(* IEC 61131-3 sources: canworks/test/plc_modbus, 6 files *)

(* ---- bridge_model.st ---- *)
(*
 * The bridge's control block and SDO registers for the block tests
 * (test/plc_modbus/run.sh), working on the blocks' LINK words directly
 * (library/modbus: 0-3 status, 4-6 control, 7-13 SDO request, 14-20 SDO
 * response): one call is one Modbus poll round. Mirrors ControlBlock and
 * SdoBridgeRegisters in plugin/src/bridge/bridge_blocks.cpp: a request runs
 * when its counter changes, the response echoes the counter. A read answers
 * 16#123456nn (nn the node); SILENT_NODE stays busy, ABORT_NODE aborts with
 * 16#06020000, writes without ALLOW_WRITE abort with 16#08000020;
 * RESTARTED answers as a bridge that just started with the request in place
 * (control result 6, SDO abort 16#08000021).
 * STruC++'s test runner does not copy a source block's in-out back, so a
 * test writes `link := bridge.LINK;` after each call.
 *)
FUNCTION_BLOCK BridgeModel
VAR_INPUT
  ALLOW_WRITE : BOOL := TRUE;
  SILENT_NODE : USINT := 99;
  ABORT_NODE : USINT := 98;
  REFUSE : BOOL;
  RESTARTED : BOOL;
END_VAR
VAR_OUTPUT
  LAST_CMD : WORD;
  LAST_NET : WORD;
  LAST_NODE : WORD;
  WRITTEN : UDINT;
  WRITTEN_SIZE : WORD;
  REQUESTS : INT;
  CONTROLS : INT;
END_VAR
VAR_IN_OUT
  LINK : ARRAY[0..1279] OF WORD;
END_VAR
VAR
  cmd : WORD;
  node : WORD;
END_VAR
  IF LINK[4] <> LINK[2] THEN
    LINK[2] := LINK[4];
    CONTROLS := CONTROLS + 1;
    LAST_CMD := SHR(LINK[5], 8);
    LAST_NET := LINK[5] AND 16#00FF;
    LAST_NODE := SHR(LINK[6], 8);
    IF RESTARTED THEN
      LINK[3] := 16#0600;
    ELSIF REFUSE THEN
      LINK[3] := 16#0500;
    ELSIF LAST_NET > 0 THEN
      LINK[3] := 16#0200;
    ELSE
      LINK[3] := 0;
    END_IF;
  END_IF;
  IF LINK[7] <> LINK[14] THEN
    LINK[14] := LINK[7];
    REQUESTS := REQUESTS + 1;
    cmd := SHR(LINK[8], 8);
    node := SHR(LINK[9], 8);
    LINK[16] := 0;
    LINK[17] := 0;
    LINK[18] := 0;
    LINK[19] := 0;
    IF RESTARTED THEN
      LINK[15] := 16#0300;
      LINK[16] := 16#0800;
      LINK[17] := 16#0021;
    ELSIF cmd = 2 AND NOT ALLOW_WRITE THEN
      LINK[15] := 16#0300;
      LINK[16] := 16#0800;
      LINK[17] := 16#0020;
    ELSIF node = USINT_TO_WORD(SILENT_NODE) THEN
      LINK[15] := 16#0100;
    ELSIF node = USINT_TO_WORD(ABORT_NODE) THEN
      LINK[15] := 16#0300;
      LINK[16] := 16#0602;
    ELSE
      LINK[15] := 16#0200;
      IF cmd = 1 THEN
        LINK[18] := 16#1234;
        LINK[19] := 16#5600 OR node;
      ELSE
        WRITTEN := DWORD_TO_UDINT(SHL(WORD_TO_DWORD(LINK[12]), 16) OR WORD_TO_DWORD(LINK[13]));
        WRITTEN_SIZE := SHR(LINK[11], 8);
      END_IF;
    END_IF;
  END_IF;
END_FUNCTION_BLOCK

(* ---- mailbox_model.st ---- *)
(*
 * The bridge's mailboxes for the block tests (test/plc_modbus/run.sh),
 * working on the blocks' LINK words directly (the places CW_LINK_SERVICE
 * describes): one call is one Modbus poll round of the bridge. Mirrors
 * plugin/src/bridge/mailboxes.cpp: a request runs when its counter changes
 * (an operation answers busy for one round, then done), the response echoes
 * the counter; STAGE and FETCH move data in 128-byte parts; receivers get
 * records in batches the program acknowledges; info and the cyclic table
 * are refreshed every round. Networks 0 and 1 exist. The bus is a set of
 * fixed answers:
 *   SDO node 98 aborts with 16#06020000, node 99 times out (2); 0x1008 the
 *   text "Valve block 24 V", 0x2000 600 bytes (byte i = i MOD 251), 0x2001
 *   300 bytes 'A' without a NUL, 0x6000 REAL32 1.5, 0x6001 REAL64 -2.25,
 *   0x6002 5 bytes, any other 16#12345600 + node (4 bytes);
 *   J1939 requests: PGN 65282 answers 40 bytes (i + 1), 65000 300 bytes
 *   (i MOD 256), 59999 a NACK (12, ACK_CODE 1), others 8 bytes (i);
 *   DM1/DM2 of any source but 77 (13): lamps 16#44, flash 16#04, codes
 *   16#00012304 and 16#0005A1FF, age 1500 ms;
 *   FIND_ECU knows one ECU, NAME 16#A00000000000ABCD at 16#33.
 * Messages come in with INJ_CAN, INJ_J1939, INJ_EMCY (INJ_RESTART: a new
 * CANopen session record); HOLD keeps them waiting for one batch; CLOSE_SLOT
 * closes a receiver as a stall would.
 * STruC++'s test runner does not copy a source block's in-out back, so a
 * test writes `link := bridge.LINK;` after each call.
 *)
FUNCTION_BLOCK MailboxModel
VAR_INPUT
  INJ_CAN : BOOL;
  INJ_J1939 : BOOL;
  INJ_EMCY : BOOL;
  INJ_RESTART : BOOL;
  INJ_ID : UDINT;
  INJ_EXT : BOOL;
  INJ_DLC : USINT := 8;
  INJ_LEN : UINT := 8;
  INJ_SRC : USINT;
  INJ_NODE : USINT;
  INJ_CODE : WORD;
  INJ_B0 : BYTE;
  CLOSE_SLOT : INT := -1;
  NO_J1939 : BOOL;
  HOLD : BOOL;           (* no new batch this round *)
  SKIP_MS : WORD;        (* extra milliseconds on the bridge's clock this round *)
  RX_BLOCKS : INT := 1;  (* receive_blocks: 95 record words, 215 with 2 *)
END_VAR
VAR_OUTPUT
  TX_COUNT : INT;
  TX_ID : UDINT;
  TX_DLC : WORD;
  TX_FLAGS : WORD;
  TX_B0 : BYTE;
  STAGES : INT;
  FETCHES : INT;
  REQUESTS : INT;
  W_LEN : UINT;
  W_KIND : WORD;
  W_SIZE : WORD;
  W_INDEX : WORD;
  J_PGN : UDINT;
  J_DEST : WORD;
  J_PRIO : WORD;
  J_LEN : UINT;
  J_COUNT : INT;
  DM_CLEARED : WORD;
  CYC_SETS : INT;
  CYC_STOPS : INT;
  STALLS : INT;
  OPEN_RX : INT;
END_VAR
VAR_IN_OUT
  LINK : ARRAY[0..1279] OF WORD;
END_VAR
VAR
  tick : WORD := 16#1000;
  seen : ARRAY[0..3] OF WORD;
  busy : ARRAY[0..3] OF INT;      (* rounds left before a running operation ends *)
  staged : ARRAY[0..7139] OF BYTE;
  staged_len : ARRAY[0..3] OF UINT;
  result : ARRAY[0..7139] OF BYTE;
  result_len : ARRAY[0..3] OF UINT;
  w_data : ARRAY[0..1784] OF BYTE;
  j_data : ARRAY[0..1784] OF BYTE;
  r : ARRAY[0..23] OF WORD;          (* results of the 4 mailboxes, 6 each *)
  st : ARRAY[0..3] OF WORD;          (* state << 8 | error *)
  rx_on : ARRAY[0..31] OF BOOL;
  rx_kind : ARRAY[0..31] OF WORD;
  rx_id : ARRAY[0..31] OF UDINT;
  rx_mask : ARRAY[0..31] OF UDINT;
  rx_flags : ARRAY[0..31] OF WORD;
  rx_gen : ARRAY[0..31] OF WORD;
  rx_drop : ARRAY[0..31] OF WORD;
  next_gen : WORD := 1;
  held : ARRAY[0..1784] OF BYTE;
  held_len : UINT;
  held_slot : INT := -1;
  (* Waiting records: receiver, kind, id/PGN/node, length, first byte, source, code, flags. *)
  q_n : INT;
  q_slot : ARRAY[0..63] OF INT;
  q_kind : ARRAY[0..63] OF WORD;
  q_id : ARRAY[0..63] OF UDINT;
  q_len : ARRAY[0..63] OF UINT;
  q_b0 : ARRAY[0..63] OF BYTE;
  q_src : ARRAY[0..63] OF WORD;
  q_code : ARRAY[0..63] OF WORD;
  q_flags : ARRAY[0..63] OF WORD;
  q_ext : ARRAY[0..63] OF BOOL;
  seq : WORD := 16#4000;
  present : DWORD;
  used : INT;
  acked : BOOL := TRUE;
  shown_rounds : INT;
  words : ARRAY[0..214] OF WORD;
  job_on : ARRAY[0..15] OF BOOL;
  job_gen : ARRAY[0..15] OF WORD;
  job_count : ARRAY[0..15] OF UDINT;
  job_keep : ARRAY[0..15] OF WORD;
  job_idle : ARRAY[0..15] OF INT;
  job_data : ARRAY[0..15] OF WORD;
  info_count : WORD;
  m : INT;
  n : INT;
  i : INT;
  k : INT;
  b : INT;
  op : WORD;
  net : WORD;
  len : UINT;
  slot : INT;
  jobs : INT;
  pending : DWORD;
  taken_long : DWORD;
  size : INT;
  room : BOOL;
  batch_tick : WORD;     (* the batch time's low word *)
  bits : DWORD;
END_VAR
  tick := tick + 10 + SKIP_MS;
  n := WORD_TO_INT(LINK[89] AND 16#0007);
  jobs := WORD_TO_INT(SHR(LINK[89], 8) AND 16#001F);
  (* ---- messages arriving on the bus ---- *)
  FOR slot := 0 TO 31 DO
    IF rx_on[slot] AND q_n < 64 THEN
      room := FALSE;
      IF INJ_CAN AND rx_kind[slot] = 1 AND (INJ_ID AND rx_mask[slot]) = (rx_id[slot] AND rx_mask[slot])
         AND INJ_EXT = ((rx_flags[slot] AND 16#0001) <> 0) THEN
        room := TRUE;
        q_kind[q_n] := 1;
        q_id[q_n] := INJ_ID;
        q_len[q_n] := USINT_TO_UINT(INJ_DLC);
      ELSIF INJ_J1939 AND rx_kind[slot] = 2 AND ((rx_flags[slot] AND 16#0001) <> 0 OR INJ_ID = rx_id[slot])
            AND (rx_mask[slot] = 255 OR USINT_TO_UDINT(INJ_SRC) = rx_mask[slot]) THEN
        room := TRUE;
        q_kind[q_n] := 2;
        q_id[q_n] := INJ_ID;
        q_len[q_n] := INJ_LEN;
      ELSIF (INJ_EMCY OR INJ_RESTART) AND rx_kind[slot] = 3 AND (rx_mask[slot] = 0 OR USINT_TO_UDINT(INJ_NODE) = rx_mask[slot]) THEN
        room := TRUE;
        q_kind[q_n] := 3;
        q_id[q_n] := USINT_TO_UDINT(INJ_NODE);
        q_len[q_n] := 5;
      END_IF;
      IF room THEN
        q_slot[q_n] := slot;
        q_b0[q_n] := INJ_B0;
        q_src[q_n] := USINT_TO_WORD(INJ_SRC);
        q_code[q_n] := INJ_CODE;
        q_ext[q_n] := INJ_EXT;
        q_flags[q_n] := SEL(INJ_RESTART, WORD#0, WORD#2);
        q_n := q_n + 1;
      END_IF;
    END_IF;
  END_FOR;
  IF CLOSE_SLOT >= 0 AND CLOSE_SLOT < 32 THEN
    rx_on[CLOSE_SLOT] := FALSE;
    present := present AND NOT SHL(DWORD#1, CLOSE_SLOT);
  END_IF;
  (* One message per call that asks for it: the inputs keep their values. *)
  INJ_CAN := FALSE;
  INJ_J1939 := FALSE;
  INJ_EMCY := FALSE;
  INJ_RESTART := FALSE;
  CLOSE_SLOT := -1;
  (* ---- request mailboxes ---- *)
  FOR m := 0 TO n - 1 DO
    b := 144 + 144 * m;
    IF busy[m] > 0 THEN
      busy[m] := busy[m] - 1;
      IF busy[m] = 0 THEN
        st[m] := SHL(WORD#2, 8) OR (st[m] AND 16#00FF);
        IF (st[m] AND 16#00FF) <> 0 THEN
          st[m] := SHL(WORD#3, 8) OR (st[m] AND 16#00FF);
        END_IF;
      END_IF;
    ELSIF LINK[b] <> seen[m] THEN
      seen[m] := LINK[b];
      REQUESTS := REQUESTS + 1;
      op := SHR(LINK[b + 1], 8);
      net := LINK[b + 1] AND 16#00FF;
      FOR i := 0 TO 5 DO
        r[6 * m + i] := 0;
      END_FOR;
      st[m] := SHL(WORD#2, 8);
      IF op = 0 THEN
        st[m] := 0;
      ELSIF op = 1 THEN
        (* STAGE *)
        STAGES := STAGES + 1;
        k := WORD_TO_INT(LINK[b + 2]);
        len := WORD_TO_UINT(LINK[b + 3]);
        FOR i := 0 TO UINT_TO_INT(len) - 1 DO
          staged[1785 * m + k + i] := WORD_TO_BYTE(SHR(LINK[b + 8 + i / 2], 8 * (1 - i MOD 2)));
        END_FOR;
        IF UINT_TO_INT(staged_len[m]) < k + UINT_TO_INT(len) THEN
          staged_len[m] := INT_TO_UINT(k + UINT_TO_INT(len));
        END_IF;
      ELSIF op = 2 THEN
        (* FETCH *)
        FETCHES := FETCHES + 1;
        k := WORD_TO_INT(LINK[b + 2]);
        r[6 * m] := UINT_TO_WORD(result_len[m]);
        FOR i := 0 TO 127 DO
          IF k + i < UINT_TO_INT(result_len[m]) THEN
            bits := BYTE_TO_DWORD(result[1785 * m + k + i]);
          ELSE
            bits := 0;
          END_IF;
          IF i MOD 2 = 0 THEN
            LINK[b + 80 + i / 2] := SHL(DWORD_TO_WORD(bits), 8);
          ELSE
            LINK[b + 80 + i / 2] := LINK[b + 80 + i / 2] OR DWORD_TO_WORD(bits);
          END_IF;
        END_FOR;
      ELSIF net > 1 AND op <> 9 AND op <> 7 THEN
        st[m] := SHL(WORD#3, 8) OR SEL(op = 3 OR op = 4, WORD#2, WORD#6);
      ELSE
        result_len[m] := 0;
        CASE WORD_TO_INT(op) OF
          3: (* SDO_READ *)
            k := WORD_TO_INT(SHR(LINK[b + 2], 8));
            busy[m] := 1;
            IF k = 98 THEN
              st[m] := 1;
              r[6 * m + 2] := 16#0602;
            ELSIF k = 99 THEN
              st[m] := 2;
              r[6 * m + 2] := 16#0504;
              busy[m] := 3;
            ELSIF LINK[b + 3] = 16#1008 THEN
              len := 16;
              FOR i := 0 TO 15 DO
                result[1785 * m + i] := 32;
              END_FOR;
              result[1785 * m] := 86;  result[1785 * m + 1] := 97;  result[1785 * m + 2] := 108;
              result[1785 * m + 3] := 118; result[1785 * m + 4] := 101; result[1785 * m + 6] := 98;
              result[1785 * m + 7] := 108; result[1785 * m + 8] := 111; result[1785 * m + 9] := 99;
              result[1785 * m + 10] := 107; result[1785 * m + 12] := 50; result[1785 * m + 13] := 52;
              result[1785 * m + 15] := 86;
            ELSIF LINK[b + 3] = 16#2000 THEN
              len := 600;
              FOR i := 0 TO 599 DO
                result[1785 * m + i] := INT_TO_BYTE(i MOD 251);
              END_FOR;
            ELSIF LINK[b + 3] = 16#2001 THEN
              len := 300;
              FOR i := 0 TO 299 DO
                result[1785 * m + i] := 65;
              END_FOR;
            ELSIF LINK[b + 3] = 16#6000 THEN
              len := 4;
              result[1785 * m] := 0; result[1785 * m + 1] := 0;
              result[1785 * m + 2] := 16#C0; result[1785 * m + 3] := 16#3F;
            ELSIF LINK[b + 3] = 16#6001 THEN
              len := 8;
              FOR i := 0 TO 5 DO
                result[1785 * m + i] := 0;
              END_FOR;
              result[1785 * m + 6] := 16#02; result[1785 * m + 7] := 16#C0;
            ELSIF LINK[b + 3] = 16#6002 THEN
              len := 5;
            ELSE
              len := 4;
              result[1785 * m] := INT_TO_BYTE(k);
              result[1785 * m + 1] := 16#56;
              result[1785 * m + 2] := 16#34;
              result[1785 * m + 3] := 16#12;
            END_IF;
            IF (st[m] AND 16#00FF) = 0 THEN
              result_len[m] := len;
              r[6 * m + 1] := UINT_TO_WORD(len);
            END_IF;
          4: (* SDO_WRITE *)
            len := WORD_TO_UINT(LINK[b + 6]);
            IF len > 128 AND staged_len[m] < len THEN
              st[m] := 6;
            ELSE
              W_LEN := len;
              W_KIND := SHR(LINK[b + 4], 8);
              W_SIZE := LINK[b + 4] AND 16#00FF;
              W_INDEX := LINK[b + 3];
              FOR i := 0 TO UINT_TO_INT(len) - 1 DO
                IF len > 128 THEN
                  w_data[i] := staged[1785 * m + i];
                ELSE
                  w_data[i] := WORD_TO_BYTE(SHR(LINK[b + 8 + i / 2], 8 * (1 - i MOD 2)));
                END_IF;
              END_FOR;
              busy[m] := 1;
            END_IF;
            staged_len[m] := 0;
          5: (* CAN_SEND *)
            TX_COUNT := TX_COUNT + 1;
            TX_ID := WORD_TO_UDINT(LINK[b + 2]) * 65536 + WORD_TO_UDINT(LINK[b + 3]);
            TX_FLAGS := SHR(LINK[b + 4], 8);
            TX_DLC := LINK[b + 4] AND 16#00FF;
            TX_B0 := WORD_TO_BYTE(SHR(LINK[b + 8], 8));
            busy[m] := 1;
          6: (* CYCLIC_SET *)
            k := WORD_TO_INT(LINK[b + 2]);
            IF jobs = 0 THEN
              st[m] := 5;
            ELSIF LINK[b + 6] = 0 OR WORD_TO_UINT(LINK[b + 6]) > 60000 THEN
              st[m] := 3;
            ELSIF LINK[b + 2] = 16#FFFF THEN
              k := -1;
              FOR i := jobs - 1 TO 0 BY -1 DO
                IF NOT job_on[i] THEN
                  k := i;
                END_IF;
              END_FOR;
              IF k < 0 THEN
                st[m] := 5;
              ELSE
                job_on[k] := TRUE;
                job_gen[k] := next_gen;
                next_gen := next_gen + 1;
                job_count[k] := 0;
                job_keep[k] := LINK[128 + k];
                job_idle[k] := 0;
                job_data[k] := LINK[b + 8];
                CYC_SETS := CYC_SETS + 1;
                r[6 * m] := INT_TO_WORD(k);
                r[6 * m + 1] := job_gen[k];
                r[6 * m + 2] := tick;
              END_IF;
            ELSIF k >= jobs OR NOT job_on[k] THEN
              st[m] := 8;
            ELSE
              job_data[k] := LINK[b + 8];
              CYC_SETS := CYC_SETS + 1;
              r[6 * m] := INT_TO_WORD(k);
              r[6 * m + 1] := job_gen[k];
              r[6 * m + 2] := tick;
            END_IF;
          7: (* CYCLIC_STOP *)
            k := WORD_TO_INT(LINK[b + 2]);
            IF k < jobs THEN
              job_on[k] := FALSE;
            END_IF;
            CYC_STOPS := CYC_STOPS + 1;
          8: (* RX_OPEN *)
            IF (LINK[89] AND 16#0010) = 0 THEN
              st[m] := 3;
            ELSE
              k := -1;
              FOR i := 31 TO 0 BY -1 DO
                IF NOT rx_on[i] THEN
                  k := i;
                END_IF;
              END_FOR;
              IF k < 0 THEN
                st[m] := 5;
              ELSE
                rx_on[k] := TRUE;
                rx_kind[k] := SHR(LINK[b + 2], 8);
                rx_flags[k] := LINK[b + 2] AND 16#00FF;
                rx_id[k] := WORD_TO_UDINT(LINK[b + 4]) * 65536 + WORD_TO_UDINT(LINK[b + 5]);
                rx_mask[k] := WORD_TO_UDINT(LINK[b + 6]) * 65536 + WORD_TO_UDINT(LINK[b + 7]);
                rx_gen[k] := next_gen;
                rx_drop[k] := 0;
                next_gen := next_gen + 1;
                r[6 * m] := INT_TO_WORD(k);
                r[6 * m + 1] := rx_gen[k];
                r[6 * m + 2] := tick;
              END_IF;
            END_IF;
          9: (* RX_CLOSE *)
            k := WORD_TO_INT(LINK[b + 2]);
            IF k < 32 THEN
              rx_on[k] := FALSE;
              present := present AND NOT SHL(DWORD#1, k);
            END_IF;
          10: (* RX_FETCH *)
            k := WORD_TO_INT(LINK[b + 2]);
            IF k <> held_slot OR NOT rx_on[k] THEN
              st[m] := 8;
            ELSE
              result_len[m] := held_len;
              FOR i := 0 TO UINT_TO_INT(held_len) - 1 DO
                result[1785 * m + i] := held[i];
              END_FOR;
              r[6 * m] := UINT_TO_WORD(held_len);
            END_IF;
          11: (* J1939_SEND *)
            len := WORD_TO_UINT(LINK[b + 5]);
            IF len > 128 AND staged_len[m] < len THEN
              st[m] := 3;
            ELSE
              J_PGN := WORD_TO_UDINT(LINK[b + 2]) * 65536 + WORD_TO_UDINT(LINK[b + 3]);
              J_DEST := SHR(LINK[b + 4], 8);
              J_PRIO := LINK[b + 4] AND 16#00FF;
              J_LEN := len;
              J_COUNT := J_COUNT + 1;
              FOR i := 0 TO UINT_TO_INT(len) - 1 DO
                IF len > 128 THEN
                  j_data[i] := staged[1785 * m + i];
                ELSE
                  j_data[i] := WORD_TO_BYTE(SHR(LINK[b + 8 + i / 2], 8 * (1 - i MOD 2)));
                END_IF;
              END_FOR;
              busy[m] := 1;
            END_IF;
            staged_len[m] := 0;
          12: (* J1939_REQUEST *)
            bits := WORD_TO_DWORD(LINK[b + 2]) * 65536 + WORD_TO_DWORD(LINK[b + 3]);
            busy[m] := 1;
            IF bits = 59999 THEN
              st[m] := 12;
              r[6 * m + 2] := 1;
            ELSE
              IF bits = 65282 THEN
                len := 40;
              ELSIF bits = 65000 THEN
                len := 300;
              ELSE
                len := 8;
              END_IF;
              FOR i := 0 TO UINT_TO_INT(len) - 1 DO
                IF bits = 65282 THEN
                  result[1785 * m + i] := INT_TO_BYTE(i + 1);
                ELSE
                  result[1785 * m + i] := INT_TO_BYTE(i MOD 256);
                END_IF;
              END_FOR;
              result_len[m] := len;
              r[6 * m] := SEL(LINK[b + 4] < 254, WORD#16#21, LINK[b + 4]);
              r[6 * m + 1] := UINT_TO_WORD(len);
            END_IF;
          13: (* DM_READ *)
            busy[m] := 1;
            IF LINK[b + 2] = 77 THEN
              st[m] := 13;
            ELSE
              r[6 * m] := 16#4404;
              r[6 * m + 1] := 2;
              r[6 * m + 3] := 1500;
              result_len[m] := 128;
              FOR i := 0 TO 127 DO
                result[1785 * m + i] := 0;
              END_FOR;
              result[1785 * m + 1] := 16#01; result[1785 * m + 2] := 16#23; result[1785 * m + 3] := 16#04;
              result[1785 * m + 5] := 16#05; result[1785 * m + 6] := 16#A1; result[1785 * m + 7] := 16#FF;
            END_IF;
          14: (* DM_CLEAR *)
            DM_CLEARED := LINK[b + 2];
            busy[m] := 1;
          15: (* FIND_ECU: NAME 16#A00000000000ABCD at 16#33 *)
            bits := 0;
            FOR i := 0 TO 3 DO
              (* (NAME xor known) and MASK, word by word *)
              bits := bits OR WORD_TO_DWORD((LINK[b + 8 + i] XOR SEL(i = 0, SEL(i = 3, WORD#0, WORD#16#ABCD), WORD#16#A000))
                                            AND LINK[b + 12 + i]);
            END_FOR;
            IF bits = 0 THEN
              r[6 * m] := 1;
              r[6 * m + 1] := 16#33;
              r[6 * m + 2] := 1;
              result_len[m] := 8;
              result[1785 * m] := 16#A0;
              FOR i := 1 TO 5 DO
                result[1785 * m + i] := 0;
              END_FOR;
              result[1785 * m + 6] := 16#AB;
              result[1785 * m + 7] := 16#CD;
            END_IF;
        ELSE
          st[m] := 3;
        END_CASE;
        IF busy[m] > 0 THEN
          (* busy now, the answer (st) shows when busy runs out *)
          st[m] := SHL(WORD#1, 8) OR (st[m] AND 16#00FF);
        ELSIF (st[m] AND 16#00FF) <> 0 THEN
          st[m] := SHL(WORD#3, 8) OR (st[m] AND 16#00FF);
        END_IF;
        IF op <> 10 THEN
          FOR i := 0 TO 127 DO
            IF i < UINT_TO_INT(result_len[m]) THEN
              bits := BYTE_TO_DWORD(result[1785 * m + i]);
            ELSE
              bits := 0;
            END_IF;
            IF i MOD 2 = 0 THEN
              LINK[b + 80 + i / 2] := SHL(DWORD_TO_WORD(bits), 8);
            ELSE
              LINK[b + 80 + i / 2] := LINK[b + 80 + i / 2] OR DWORD_TO_WORD(bits);
            END_IF;
          END_FOR;
        ELSE
          FOR i := 0 TO 127 DO
            IF i < UINT_TO_INT(held_len) THEN
              bits := BYTE_TO_DWORD(held[i]);
            ELSE
              bits := 0;
            END_IF;
            IF i MOD 2 = 0 THEN
              LINK[b + 80 + i / 2] := SHL(DWORD_TO_WORD(bits), 8);
            ELSE
              LINK[b + 80 + i / 2] := LINK[b + 80 + i / 2] OR DWORD_TO_WORD(bits);
            END_IF;
          END_FOR;
        END_IF;
      END_IF;
    END_IF;
    (* the response *)
    LINK[b + 72] := seen[m];
    LINK[b + 73] := st[m];
    IF SHR(st[m], 8) = 1 THEN
      FOR i := 0 TO 5 DO
        LINK[b + 74 + i] := 0;
      END_FOR;
    ELSE
      FOR i := 0 TO 5 DO
        LINK[b + 74 + i] := r[6 * m + i];
      END_FOR;
    END_IF;
  END_FOR;
  (* ---- receive mailbox ---- *)
  IF (LINK[89] AND 16#0010) <> 0 THEN
    IF NOT acked THEN
      pending := SHL(WORD_TO_DWORD(LINK[103]), 16) OR WORD_TO_DWORD(LINK[104]);
      IF LINK[102] = seq AND (pending AND present) = 0 THEN
        acked := TRUE;
      ELSE
        shown_rounds := shown_rounds + 1;
        IF shown_rounds >= 100 THEN
          (* the stall rule: close the receivers that kept the batch *)
          FOR i := 0 TO 31 DO
            IF (SHR(present, i) AND 1) <> 0 AND (LINK[102] <> seq OR (SHR(pending, i) AND 1) <> 0) THEN
              rx_on[i] := FALSE;
            END_IF;
          END_FOR;
          STALLS := STALLS + 1;
          acked := TRUE;
        END_IF;
      END_IF;
    END_IF;
    IF acked AND q_n > 0 AND NOT HOLD THEN
      used := 0;
      present := 0;
      taken_long := 0;
      k := 0;
      (* records in arrival order while they fit; one long J1939 per receiver *)
      WHILE k < q_n DO
        slot := q_slot[k];
        size := 7;
        IF q_kind[k] = 1 THEN
          size := 10;
        ELSIF q_kind[k] = 2 THEN
          size := 12;
        ELSIF q_kind[k] = 3 THEN
          size := 12;
        END_IF;
        IF NOT rx_on[slot] THEN
          (* closed: its records go *)
          FOR i := k TO q_n - 2 DO
            q_slot[i] := q_slot[i + 1]; q_kind[i] := q_kind[i + 1]; q_id[i] := q_id[i + 1];
            q_len[i] := q_len[i + 1]; q_b0[i] := q_b0[i + 1]; q_src[i] := q_src[i + 1];
            q_code[i] := q_code[i + 1]; q_flags[i] := q_flags[i + 1]; q_ext[i] := q_ext[i + 1];
          END_FOR;
          q_n := q_n - 1;
        ELSIF used + size > SEL(RX_BLOCKS = 2, 95, 215) OR (SHR(taken_long, slot) AND 1) <> 0 THEN
          k := q_n;
        ELSE
          words[used] := SHL(INT_TO_WORD(slot), 8) OR SHL(q_kind[k], 4) OR q_flags[k];
          words[used + 1] := 0;
          FOR i := k + 1 TO q_n - 1 DO
            IF q_slot[i] = slot THEN
              words[used + 1] := words[used + 1] + 1;
            END_IF;
          END_FOR;
          words[used + 2] := rx_drop[slot];
          IF q_kind[k] = 1 THEN
            words[used + 3] := UDINT_TO_WORD(SHR(q_id[k], 16));
            words[used + 4] := UDINT_TO_WORD(q_id[k]);
            words[used + 5] := SEL(q_ext[k], WORD#0, WORD#16#0100) OR UINT_TO_WORD(q_len[k]);
            FOR i := 0 TO 3 DO
              words[used + 6 + i] := SHL(BYTE_TO_WORD(q_b0[k]) + INT_TO_WORD(2 * i), 8) OR
                                      ((BYTE_TO_WORD(q_b0[k]) + INT_TO_WORD(2 * i + 1)) AND 16#00FF);
            END_FOR;
          ELSIF q_kind[k] = 2 THEN
            words[used + 3] := UDINT_TO_WORD(SHR(q_id[k], 16));
            words[used + 4] := UDINT_TO_WORD(q_id[k]);
            words[used + 5] := SHL(q_src[k], 8) OR 16#00FF;
            words[used + 6] := 6;
            words[used + 7] := UINT_TO_WORD(q_len[k]);
            FOR i := 0 TO 3 DO
              words[used + 8 + i] := SHL(BYTE_TO_WORD(q_b0[k]) + INT_TO_WORD(2 * i), 8) OR
                                      ((BYTE_TO_WORD(q_b0[k]) + INT_TO_WORD(2 * i + 1)) AND 16#00FF);
            END_FOR;
            IF q_len[k] > 8 THEN
              words[used] := words[used] OR 16#0001;
              taken_long := taken_long OR SHL(DWORD#1, slot);
              held_slot := slot;
              held_len := q_len[k];
              FOR i := 0 TO UINT_TO_INT(q_len[k]) - 1 DO
                held[i] := INT_TO_BYTE((BYTE_TO_INT(q_b0[k]) + i) MOD 256);
              END_FOR;
            END_IF;
          ELSE
            words[used + 3] := 0;
            words[used + 4] := 16#0006;
            words[used + 5] := 16#0000;
            words[used + 6] := tick;
            words[used + 7] := SHL(UDINT_TO_WORD(q_id[k]), 8) OR 16#0081;
            words[used + 8] := q_code[k];
            words[used + 9] := 16#0102;
            words[used + 10] := 16#0304;
            words[used + 11] := 16#0500;
          END_IF;
          used := used + size;
          present := present OR SHL(DWORD#1, slot);
          FOR i := k TO q_n - 2 DO
            q_slot[i] := q_slot[i + 1]; q_kind[i] := q_kind[i + 1]; q_id[i] := q_id[i + 1];
            q_len[i] := q_len[i + 1]; q_b0[i] := q_b0[i + 1]; q_src[i] := q_src[i + 1];
            q_code[i] := q_code[i + 1]; q_flags[i] := q_flags[i + 1]; q_ext[i] := q_ext[i + 1];
          END_FOR;
          q_n := q_n - 1;
        END_IF;
      END_WHILE;
      IF present <> 0 THEN
        seq := seq + 1;
        batch_tick := tick;
        acked := FALSE;
        shown_rounds := 0;
      END_IF;
    END_IF;
    LINK[720] := seq;
    LINK[721] := DWORD_TO_WORD(SHR(present, 16));
    LINK[722] := DWORD_TO_WORD(present);
    LINK[723] := INT_TO_WORD(used);
    LINK[724] := tick;
    LINK[741] := 0;
    LINK[742] := 16#0006;
    LINK[743] := 16#0000;
    LINK[744] := batch_tick;
    OPEN_RX := 0;
    FOR i := 0 TO 15 DO
      LINK[725 + i] := SHL(SEL(rx_on[2 * i], WORD#0, rx_gen[2 * i] AND 16#00FF), 8) OR
                       SEL(rx_on[2 * i + 1], WORD#0, rx_gen[2 * i + 1] AND 16#00FF);
    END_FOR;
    FOR i := 0 TO 31 DO
      IF rx_on[i] THEN
        OPEN_RX := OPEN_RX + 1;
      END_IF;
    END_FOR;
    FOR i := 0 TO SEL(RX_BLOCKS = 2, 94, 214) DO
      LINK[745 + i] := words[i];
    END_FOR;
  END_IF;
  (* ---- network info: network 0 a J1939 network, network 1 not ---- *)
  IF (LINK[89] AND 16#0020) <> 0 THEN
    info_count := info_count + 1;
    FOR k := 0 TO 1 DO
      b := 960 + 18 * k;
      LINK[b] := 16#000C;
      LINK[b + 1] := 1;
      LINK[b + 2] := 2;
      LINK[b + 3] := 0;
      LINK[b + 4] := 3;
      LINK[b + 5] := 0;
      LINK[b + 6] := 1000;
      LINK[b + 7] := 1;
      LINK[b + 8] := 0;
      LINK[b + 9] := 0;
      LINK[b + 10] := 5;
      IF k = 0 AND NOT NO_J1939 THEN
        LINK[b + 11] := 16#0180;
        LINK[b + 12] := 16#A000;
        LINK[b + 13] := 0;
        LINK[b + 14] := 0;
        LINK[b + 15] := 16#ABCD;
        LINK[b + 16] := 4;
      ELSE
        LINK[b + 11] := 16#FF0A;
        LINK[b + 12] := 0;
        LINK[b + 13] := 0;
        LINK[b + 14] := 0;
        LINK[b + 15] := 0;
        LINK[b + 16] := 0;
      END_IF;
      LINK[b + 17] := info_count;
    END_FOR;
  END_IF;
  (* ---- cyclic job table and keepalives ---- *)
  IF jobs > 0 THEN
    LINK[1104] := tick;
    FOR k := 0 TO jobs - 1 DO
      b := 1105 + 4 * k;
      IF job_on[k] THEN
        IF LINK[128 + k] = job_keep[k] THEN
          job_idle[k] := job_idle[k] + 1;
          IF job_idle[k] >= 100 THEN
            job_on[k] := FALSE;
          END_IF;
        ELSE
          job_keep[k] := LINK[128 + k];
          job_idle[k] := 0;
        END_IF;
      END_IF;
      IF job_on[k] THEN
        job_count[k] := job_count[k] + 1;
        LINK[b] := 16#0100;
        LINK[b + 1] := job_gen[k];
        LINK[b + 2] := UDINT_TO_WORD(SHR(job_count[k], 16));
        LINK[b + 3] := UDINT_TO_WORD(job_count[k]);
      ELSE
        LINK[b] := 0;
        LINK[b + 1] := 0;
        LINK[b + 2] := 0;
        LINK[b + 3] := 0;
      END_IF;
    END_FOR;
  END_IF;
END_FUNCTION_BLOCK

(* ---- test_bits.st ---- *)
(*
 * Bit channels of PDO entries on the bridge (canopen-pdo-io "Bit channels in
 * the generated programs on the bridge"): the generated canworks_in and
 * canworks_out for examples/openplc-modbus with bits on rtd TPDO1 0x7130:1
 * (bit 9), dio TPDO1 0x6000:1 (bits 0 and 3) and dio RPDO1 0x6200:1 (bit 2),
 * as function blocks (make_programs.py, bits.st). Run by test/plc_modbus/run.sh.
 *)
TEST 'canworks_in reads each bit from its entry'
  VAR
    cin : canworks_in_fb;
  END_VAR
  cin.i6 := 16#0200;
  cin.i10 := 16#0900;
  cin();
  ASSERT_TRUE(cin.canworks.rtd_hi);
  ASSERT_EQ(cin.canworks.rtd_AI0_Input_PV, 512);
  ASSERT_TRUE(cin.canworks.dio_first_bit);
  ASSERT_TRUE(cin.canworks.dio_Read_input_8_bit_1_bit3);
  ASSERT_EQ(cin.canworks.dio_Read_input_8_bit_1, 9);
  cin.i6 := 16#01FF;
  cin.i10 := 16#F6FF;
  cin();
  ASSERT_FALSE(cin.canworks.rtd_hi);
  ASSERT_FALSE(cin.canworks.dio_first_bit);
  ASSERT_FALSE(cin.canworks.dio_Read_input_8_bit_1_bit3);
END_TEST

TEST 'canworks_out ORs each bit into its entry word'
  VAR
    cout : canworks_out_fb;
  END_VAR
  cout.canworks.dio_Write_output_8_bit_1 := 16#01;
  cout.canworks.dio_Write_output_8_bit_2 := 16#22;
  cout();
  ASSERT_EQ(cout.q3, 16#0122);
  cout.canworks.dio_lamp := TRUE;
  cout();
  ASSERT_EQ(cout.q3, 16#0522);
  cout.canworks.dio_Write_output_8_bit_1 := 0;
  cout();
  ASSERT_EQ(cout.q3, 16#0422);
END_TEST

(* ---- test_blocks.st ---- *)
(*
 * The canworks blocks over the bridge (library/modbus) against the bridge
 * model. LINK word 21 holds the flags: 16#0001 the bridge answers, 16#0002
 * a control block, 16#0004 SDO registers, 16#0100 << n a live list for
 * network n. Run by test/plc_modbus/run.sh.
 *)
TEST 'SDO read through the bridge registers'
  VAR
    link : ARRAY[0..1279] OF WORD;
    bridge : BridgeModel;
    rd : CO_SDO_READ;
  END_VAR
  link[21] := 16#0005;
  rd(EXECUTE := TRUE, NODE := 5, INDEX := 16#1018, SUBINDEX := 1, LINK := link);
  ASSERT_TRUE(rd.BUSY);
  ASSERT_EQ(link[8], 16#0100);
  ASSERT_EQ(link[9], 16#0501);
  ASSERT_EQ(link[10], 16#1018);
  bridge(LINK := link);
  link := bridge.LINK;
  rd(EXECUTE := TRUE, NODE := 5, INDEX := 16#1018, SUBINDEX := 1, LINK := link);
  ASSERT_TRUE(rd.DONE);
  ASSERT_FALSE(rd.BUSY);
  ASSERT_EQ(rd.DATA, 16#12345605);
  ASSERT_EQ(link[23], 0);
  rd(EXECUTE := TRUE, NODE := 5, INDEX := 16#1018, SUBINDEX := 1, LINK := link);
  ASSERT_TRUE(rd.DONE);
  rd(EXECUTE := FALSE, NODE := 5, INDEX := 16#1018, SUBINDEX := 1, LINK := link);
  ASSERT_FALSE(rd.DONE);
END_TEST

TEST 'two instances in one scan share the SDO registers'
  VAR
    link : ARRAY[0..1279] OF WORD;
    bridge : BridgeModel;
    r1 : CO_SDO_READ;
    r2 : CO_SDO_READ;
    i : INT;
  END_VAR
  link[21] := 16#0005;
  r1(EXECUTE := TRUE, NODE := 5, INDEX := 16#1000, LINK := link);
  r2(EXECUTE := TRUE, NODE := 6, INDEX := 16#1000, LINK := link);
  ASSERT_TRUE(r2.BUSY);
  ASSERT_EQ(link[23], r1.me);
  bridge(LINK := link);
  link := bridge.LINK;
  FOR i := 1 TO 5 DO
    r1(EXECUTE := TRUE, NODE := 5, INDEX := 16#1000, LINK := link);
    r2(EXECUTE := TRUE, NODE := 6, INDEX := 16#1000, LINK := link);
    bridge(LINK := link);
    link := bridge.LINK;
  END_FOR;
  ASSERT_TRUE(r1.DONE);
  ASSERT_TRUE(r2.DONE);
  ASSERT_EQ(r1.DATA, 16#12345605);
  ASSERT_EQ(r2.DATA, 16#12345606);
  ASSERT_EQ(bridge.REQUESTS, 2);
END_TEST

TEST 'SDO write sends the value and size'
  VAR
    link : ARRAY[0..1279] OF WORD;
    bridge : BridgeModel;
    wr : CO_SDO_WRITE;
  END_VAR
  link[21] := 16#0005;
  wr(EXECUTE := TRUE, NODE := 7, INDEX := 16#2000, SUBINDEX := 3, DATA := 16#AABBCCDD, SIZE := 4, LINK := link);
  bridge(LINK := link);
  link := bridge.LINK;
  wr(EXECUTE := TRUE, NODE := 7, INDEX := 16#2000, SUBINDEX := 3, DATA := 16#AABBCCDD, SIZE := 4, LINK := link);
  ASSERT_TRUE(wr.DONE);
  ASSERT_EQ(bridge.WRITTEN, 16#AABBCCDD);
  ASSERT_EQ(bridge.WRITTEN_SIZE, 4);
END_TEST

TEST 'bridge not reachable ends at once with 20'
  VAR
    link : ARRAY[0..1279] OF WORD;
    rd : CO_SDO_READ;
    nmt : CO_NMT;
  END_VAR
  link[21] := 16#0006;
  rd(EXECUTE := TRUE, NODE := 5, LINK := link);
  ASSERT_TRUE(rd.ERROR);
  ASSERT_FALSE(rd.BUSY);
  ASSERT_EQ(rd.ERROR_ID, 20);
  nmt(EXECUTE := TRUE, NODE := 5, COMMAND := 1, LINK := link);
  ASSERT_EQ(nmt.ERROR_ID, 20);
END_TEST

TEST 'link lost while busy ends with 20 and frees the registers'
  VAR
    link : ARRAY[0..1279] OF WORD;
    bridge : BridgeModel;
    rd : CO_SDO_READ;
  END_VAR
  link[21] := 16#0005;
  bridge.SILENT_NODE := 9;
  rd(EXECUTE := TRUE, NODE := 9, LINK := link);
  bridge(LINK := link);
  link := bridge.LINK;
  link[21] := 16#0004;
  rd(EXECUTE := TRUE, NODE := 9, LINK := link);
  ASSERT_EQ(rd.ERROR_ID, 20);
  ASSERT_EQ(link[23], 0);
END_TEST

TEST 'writes not allowed by the config end with 21'
  VAR
    link : ARRAY[0..1279] OF WORD;
    bridge : BridgeModel;
    wr : CO_SDO_WRITE;
  END_VAR
  link[21] := 16#0005;
  bridge.ALLOW_WRITE := FALSE;
  wr(EXECUTE := TRUE, NODE := 7, INDEX := 16#2000, DATA := 1, SIZE := 1, LINK := link);
  bridge(LINK := link);
  link := bridge.LINK;
  wr(EXECUTE := TRUE, NODE := 7, INDEX := 16#2000, DATA := 1, SIZE := 1, LINK := link);
  ASSERT_TRUE(wr.ERROR);
  ASSERT_EQ(wr.ERROR_ID, 21);
  ASSERT_EQ(wr.ABORT_CODE, 16#08000020);
END_TEST

TEST 'a request the restarted bridge did not run ends with 8'
  VAR
    link : ARRAY[0..1279] OF WORD;
    bridge : BridgeModel;
    rd : CO_SDO_READ;
    nmt : CO_NMT;
  END_VAR
  link[21] := 16#0007;
  bridge.RESTARTED := TRUE;
  rd(EXECUTE := TRUE, NODE := 7, INDEX := 16#1018, SUBINDEX := 1, LINK := link);
  nmt(EXECUTE := TRUE, NODE := 7, COMMAND := 1, LINK := link);
  bridge(LINK := link);
  link := bridge.LINK;
  rd(EXECUTE := TRUE, NODE := 7, INDEX := 16#1018, SUBINDEX := 1, LINK := link);
  nmt(EXECUTE := TRUE, NODE := 7, COMMAND := 1, LINK := link);
  ASSERT_TRUE(rd.ERROR);
  ASSERT_EQ(rd.ERROR_ID, 8);
  ASSERT_EQ(rd.ABORT_CODE, 16#08000021);
  ASSERT_TRUE(nmt.ERROR);
  ASSERT_EQ(nmt.ERROR_ID, 8);
END_TEST

TEST 'node abort ends with 1 and the abort code'
  VAR
    link : ARRAY[0..1279] OF WORD;
    bridge : BridgeModel;
    rd : CO_SDO_READ;
  END_VAR
  link[21] := 16#0005;
  rd(EXECUTE := TRUE, NODE := 98, INDEX := 16#6000, LINK := link);
  bridge(LINK := link);
  link := bridge.LINK;
  rd(EXECUTE := TRUE, NODE := 98, INDEX := 16#6000, LINK := link);
  ASSERT_EQ(rd.ERROR_ID, 1);
  ASSERT_EQ(rd.ABORT_CODE, 16#06020000);
END_TEST

TEST 'no answer within TIMEOUT ends with 2'
  VAR
    link : ARRAY[0..1279] OF WORD;
    bridge : BridgeModel;
    rd : CO_SDO_READ;
  END_VAR
  link[21] := 16#0005;
  bridge.SILENT_NODE := 9;
  rd(EXECUTE := TRUE, NODE := 9, TIMEOUT := T#100ms, LINK := link);
  bridge(LINK := link);
  link := bridge.LINK;
  ADVANCE_TIME(T#40ms);
  rd(EXECUTE := TRUE, NODE := 9, TIMEOUT := T#100ms, LINK := link);
  bridge(LINK := link);
  link := bridge.LINK;
  ADVANCE_TIME(T#40ms);
  rd(EXECUTE := TRUE, NODE := 9, TIMEOUT := T#100ms, LINK := link);
  ASSERT_TRUE(rd.BUSY);
  ADVANCE_TIME(T#40ms);
  rd(EXECUTE := TRUE, NODE := 9, TIMEOUT := T#100ms, LINK := link);
  ASSERT_TRUE(rd.ERROR);
  ASSERT_EQ(rd.ERROR_ID, 2);
  ASSERT_EQ(link[23], 0);
END_TEST

TEST 'invalid input and missing registers'
  VAR
    link : ARRAY[0..1279] OF WORD;
    rd : CO_SDO_READ;
    wr : CO_SDO_WRITE;
    nmt : CO_NMT;
  END_VAR
  link[21] := 16#0001;
  rd(EXECUTE := TRUE, NODE := 5, LINK := link);
  ASSERT_EQ(rd.ERROR_ID, 22);
  nmt(EXECUTE := TRUE, NODE := 5, COMMAND := 1, LINK := link);
  ASSERT_EQ(nmt.ERROR_ID, 22);
  link[21] := 16#0007;
  wr(EXECUTE := TRUE, NODE := 5, SIZE := 5, LINK := link);
  ASSERT_EQ(wr.ERROR_ID, 6);
  nmt(EXECUTE := FALSE, LINK := link);
  nmt(EXECUTE := TRUE, NODE := 5, COMMAND := 3, LINK := link);
  ASSERT_EQ(nmt.ERROR_ID, 6);
END_TEST

TEST 'NMT through the control block'
  VAR
    link : ARRAY[0..1279] OF WORD;
    bridge : BridgeModel;
    nmt : CO_NMT;
  END_VAR
  link[21] := 16#0003;
  nmt(EXECUTE := TRUE, NODE := 5, COMMAND := 2, LINK := link);
  ASSERT_TRUE(nmt.BUSY);
  bridge(LINK := link);
  link := bridge.LINK;
  nmt(EXECUTE := TRUE, NODE := 5, COMMAND := 2, LINK := link);
  ASSERT_TRUE(nmt.DONE);
  ASSERT_EQ(bridge.LAST_CMD, 4);
  ASSERT_EQ(bridge.LAST_NODE, 5);
  ASSERT_EQ(link[22], 0);
  nmt(EXECUTE := FALSE, LINK := link);
  bridge.REFUSE := TRUE;
  nmt(EXECUTE := TRUE, NODE := 0, COMMAND := 128, LINK := link);
  bridge(LINK := link);
  link := bridge.LINK;
  nmt(EXECUTE := TRUE, NODE := 0, COMMAND := 128, LINK := link);
  ASSERT_EQ(nmt.ERROR_ID, 5);
  ASSERT_EQ(bridge.LAST_CMD, 5);
  ASSERT_EQ(bridge.CONTROLS, 2);
END_TEST

TEST 'node live from the live list'
  VAR
    link : ARRAY[0..1279] OF WORD;
    live : CO_NODE_LIVE;
  END_VAR
  link[21] := 16#0201;
  link[33] := 16#2002;
  live(NETWORK := 1, NODE := 5, LINK := link);
  ASSERT_TRUE(live.LIVE);
  live(NETWORK := 1, NODE := 9, LINK := link);
  ASSERT_TRUE(live.LIVE);
  live(NETWORK := 1, NODE := 6, LINK := link);
  ASSERT_FALSE(live.LIVE);
  live(NETWORK := 0, NODE := 5, LINK := link);
  ASSERT_FALSE(live.LIVE);
  link[21] := 16#0200;
  live(NETWORK := 1, NODE := 5, LINK := link);
  ASSERT_FALSE(live.LIVE);
END_TEST

TEST 'REAL and LREAL bit patterns'
  ASSERT_EQ(CW_REAL_TO_DWORD(1.0), DWORD#16#3F800000);
  ASSERT_EQ(CW_REAL_TO_DWORD(-2.5), DWORD#16#C0200000);
  ASSERT_EQ(CW_REAL_TO_DWORD(0.1), DWORD#16#3DCCCCCD);
  ASSERT_EQ(CW_REAL_TO_DWORD(0.0), DWORD#0);
  ASSERT_NEAR(CW_DWORD_TO_REAL(DWORD#16#40490FDB), 3.14159265, 0.000001);
  ASSERT_EQ(CW_REAL_TO_DWORD(CW_DWORD_TO_REAL(DWORD#16#00000001)), DWORD#16#00000001);
  ASSERT_EQ(CW_REAL_TO_DWORD(CW_DWORD_TO_REAL(DWORD#16#7F7FFFFF)), DWORD#16#7F7FFFFF);
  ASSERT_EQ(CW_REAL_TO_DWORD(CW_DWORD_TO_REAL(DWORD#16#C2F6E979)), DWORD#16#C2F6E979);
  ASSERT_EQ(CW_LREAL_TO_LWORD(-2.5), LWORD#16#C004000000000000);
  ASSERT_EQ(CW_LREAL_TO_LWORD(0.1), LWORD#16#3FB999999999999A);
  ASSERT_EQ(CW_LREAL_TO_LWORD(CW_LWORD_TO_LREAL(LWORD#16#0000000000000001)), LWORD#16#0000000000000001);
  ASSERT_EQ(CW_LREAL_TO_LWORD(CW_LWORD_TO_LREAL(LWORD#16#7FEFFFFFFFFFFFFF)), LWORD#16#7FEFFFFFFFFFFFFF);
  ASSERT_NEAR(CW_LWORD_TO_LREAL(LWORD#16#400921FB54442D18), 3.141592653589793, 0.000000000001);
END_TEST

(* ---- test_mailbox_blocks.st ---- *)
(*
 * The canworks blocks over the bridge's mailboxes (library/modbus) against
 * the mailbox model. A scan: CW_LINK_SERVICE, the blocks, then one model
 * round (one Modbus poll). LINK word 21 bit 0: the bridge answers; word 89:
 * the mailbox flags (16#0431: one request mailbox, the receive mailbox,
 * network info, 4 cyclic jobs). Run by test/plc_modbus/run.sh.
 *)
TEST 'link service counts scans, moves tickets and frees a forgotten mailbox'
  VAR
    link : ARRAY[0..1279] OF WORD;
    svc : CW_LINK_SERVICE;
    i : INT;
  END_VAR
  link[21] := 1;
  link[89] := 16#0431;
  link[92] := 7;
  link[94] := 5;
  link[98] := 0;
  svc(LINK := link);
  ASSERT_EQ(link[90], 1);
  ASSERT_EQ(link[93], 7);
  ASSERT_EQ(link[92], 0);
  FOR i := 1 TO 100 DO
    svc(LINK := link);
  END_FOR;
  ASSERT_EQ(link[94], 0);
  (* a new batch: acknowledged, its receivers pending *)
  link[720] := 16#4321;
  link[721] := 16#0001;
  link[722] := 16#0004;
  svc(LINK := link);
  ASSERT_EQ(link[102], 16#4321);
  ASSERT_EQ(link[103], 16#0001);
  ASSERT_EQ(link[104], 16#0004);
  (* bridge gone: requests and acknowledgement cleared *)
  link[21] := 0;
  link[145] := 16#0500;
  link[94] := 3;
  svc(LINK := link);
  ASSERT_EQ(link[145], 0);
  ASSERT_EQ(link[94], 0);
  ASSERT_EQ(link[102], 0);
END_TEST

TEST 'three senders share one mailbox in call order'
  VAR
    link : ARRAY[0..1279] OF WORD;
    svc : CW_LINK_SERVICE;
    bridge : MailboxModel;
    s1 : CAN_SEND;
    s2 : CAN_SEND;
    s3 : CAN_SEND;
    d : ARRAY[0..7] OF BYTE;
    i : INT;
    first2 : INT;
  END_VAR
  link[21] := 1;
  link[89] := 16#0431;
  d[0] := 16#11;
  FOR i := 1 TO 12 DO
    svc(LINK := link);
    s1(EXECUTE := TRUE, ID := 16#101, DLC := 1, DATA := d, LINK := link);
    s2(EXECUTE := TRUE, ID := 16#102, DLC := 1, DATA := d, LINK := link);
    s3(EXECUTE := TRUE, ID := 16#103, DLC := 1, DATA := d, LINK := link);
    bridge(LINK := link);
    link := bridge.LINK;
    IF bridge.TX_COUNT = 2 AND first2 = 0 THEN
      first2 := i;
      ASSERT_EQ(bridge.TX_ID, 16#102);
    END_IF;
  END_FOR;
  ASSERT_TRUE(s1.DONE);
  ASSERT_TRUE(s2.DONE);
  ASSERT_TRUE(s3.DONE);
  ASSERT_EQ(bridge.TX_COUNT, 3);
  ASSERT_EQ(bridge.TX_ID, 16#103);
  ASSERT_EQ(bridge.TX_B0, 16#11);
  ASSERT_EQ(link[94], 0);
END_TEST

TEST 'without mailboxes or bridge the blocks end in the same call'
  VAR
    link : ARRAY[0..1279] OF WORD;
    snd : CAN_SEND;
    rd : CO_SDO_READ_STRING;
    rx : CAN_RECEIVE;
    info : CAN_BUS_INFO;
    d : ARRAY[0..7] OF BYTE;
  END_VAR
  link[21] := 1;
  snd(EXECUTE := TRUE, ID := 1, DLC := 0, DATA := d, LINK := link);
  ASSERT_TRUE(snd.ERROR);
  ASSERT_EQ(snd.ERROR_ID, 22);
  rd(EXECUTE := TRUE, NODE := 5, INDEX := 16#1008, LINK := link);
  ASSERT_EQ(rd.ERROR_ID, 22);
  rx(ENABLE := TRUE, ID := 1, RX_DATA := d, LINK := link);
  ASSERT_EQ(rx.ERROR_ID, 22);
  info(NETWORK := 0, LINK := link);
  ASSERT_EQ(info.ERROR_ID, 22);
  link[21] := 0;
  link[89] := 16#0431;
  snd(EXECUTE := FALSE, DATA := d, LINK := link);
  snd(EXECUTE := TRUE, ID := 1, DLC := 9, DATA := d, LINK := link);
  ASSERT_EQ(snd.ERROR_ID, 3);
  snd(EXECUTE := FALSE, DATA := d, LINK := link);
  snd(EXECUTE := TRUE, ID := 1, DLC := 0, DATA := d, LINK := link);
  ASSERT_EQ(snd.ERROR_ID, 20);
END_TEST

TEST 'SDO string, bytes and REAL reads'
  VAR
    link : ARRAY[0..1279] OF WORD;
    svc : CW_LINK_SERVICE;
    bridge : MailboxModel;
    rs : CO_SDO_READ_STRING;
    rb : CO_SDO_READ_BYTES;
    r4 : CO_SDO_READ_REAL;
    r8 : CO_SDO_READ_REAL;
    r5 : CO_SDO_READ_REAL;
    long : CO_SDO_READ_STRING;
    buf : ARRAY[0..1023] OF BYTE;
    i : INT;
  END_VAR
  link[21] := 1;
  link[89] := 16#0431;
  FOR i := 1 TO 40 DO
    svc(LINK := link);
    rs(EXECUTE := TRUE, NODE := 5, INDEX := 16#1008, LINK := link);
    rb(EXECUTE := TRUE, NODE := 5, INDEX := 16#2000, BUFFER := buf, LINK := link);
    r4(EXECUTE := TRUE, NODE := 5, INDEX := 16#6000, LINK := link);
    r8(EXECUTE := TRUE, NODE := 5, INDEX := 16#6001, LINK := link);
    r5(EXECUTE := TRUE, NODE := 5, INDEX := 16#6002, LINK := link);
    long(EXECUTE := TRUE, NODE := 5, INDEX := 16#2001, LINK := link);
    bridge(LINK := link);
    link := bridge.LINK;
  END_FOR;
  ASSERT_TRUE(rs.DONE);
  ASSERT_EQ(rs.VALUE, 'Valve block 24 V');
  ASSERT_TRUE(rb.DONE);
  ASSERT_EQ(rb.SIZE, 600);
  ASSERT_EQ(buf[0], 0);
  ASSERT_EQ(buf[300], 49);
  ASSERT_EQ(buf[599], 97);
  ASSERT_TRUE(r4.DONE);
  ASSERT_EQ(r4.VALUE, 1.5);
  ASSERT_TRUE(r8.DONE);
  ASSERT_EQ(r8.VALUE, -2.25);
  ASSERT_TRUE(r5.ERROR);
  ASSERT_EQ(r5.ERROR_ID, 7);
  ASSERT_TRUE(long.ERROR);
  ASSERT_EQ(long.ERROR_ID, 7);
  ASSERT_EQ(bridge.FETCHES, 5);
END_TEST

TEST 'SDO writes: 600 bytes staged, a string, a REAL32'
  VAR
    link : ARRAY[0..1279] OF WORD;
    svc : CW_LINK_SERVICE;
    bridge : MailboxModel;
    wb : CO_SDO_WRITE_BYTES;
    ws : CO_SDO_WRITE_STRING;
    wr : CO_SDO_WRITE_REAL;
    buf : ARRAY[0..1023] OF BYTE;
    i : INT;
  END_VAR
  link[21] := 1;
  link[89] := 16#0431;
  FOR i := 0 TO 599 DO
    buf[i] := INT_TO_BYTE(i MOD 7);
  END_FOR;
  FOR i := 1 TO 20 DO
    svc(LINK := link);
    wb(EXECUTE := TRUE, NODE := 5, INDEX := 16#2000, SIZE := 600, BUFFER := buf, LINK := link);
    bridge(LINK := link);
    link := bridge.LINK;
  END_FOR;
  ASSERT_TRUE(wb.DONE);
  ASSERT_EQ(bridge.W_LEN, 600);
  ASSERT_EQ(bridge.w_data[599], 4);
  ASSERT_EQ(bridge.w_data[128], 2);
  ASSERT_EQ(bridge.STAGES, 5);
  FOR i := 1 TO 6 DO
    svc(LINK := link);
    ws(EXECUTE := TRUE, NODE := 5, INDEX := 16#2002, VALUE := 'abc', LINK := link);
    bridge(LINK := link);
    link := bridge.LINK;
  END_FOR;
  ASSERT_TRUE(ws.DONE);
  ASSERT_EQ(bridge.W_LEN, 3);
  ASSERT_EQ(bridge.W_KIND, 2);
  ASSERT_EQ(bridge.w_data[2], 99);
  FOR i := 1 TO 6 DO
    svc(LINK := link);
    wr(EXECUTE := TRUE, NODE := 5, INDEX := 16#6000, VALUE := 1.5, SIZE := 4, LINK := link);
    bridge(LINK := link);
    link := bridge.LINK;
  END_FOR;
  ASSERT_TRUE(wr.DONE);
  ASSERT_EQ(bridge.W_LEN, 8);
  ASSERT_EQ(bridge.W_KIND, 1);
  ASSERT_EQ(bridge.W_SIZE, 4);
  ASSERT_EQ(bridge.w_data[6], 16#F8);
  ASSERT_EQ(bridge.w_data[7], 16#3F);
END_TEST

TEST 'SDO abort and timeout keep the bridge answer'
  VAR
    link : ARRAY[0..1279] OF WORD;
    svc : CW_LINK_SERVICE;
    bridge : MailboxModel;
    ra : CO_SDO_READ_BYTES;
    rt : CO_SDO_READ_STRING;
    buf : ARRAY[0..1023] OF BYTE;
    i : INT;
  END_VAR
  link[21] := 1;
  link[89] := 16#0431;
  FOR i := 1 TO 12 DO
    svc(LINK := link);
    ra(EXECUTE := TRUE, NODE := 98, INDEX := 16#2000, BUFFER := buf, LINK := link);
    rt(EXECUTE := TRUE, NODE := 99, INDEX := 16#1008, LINK := link);
    bridge(LINK := link);
    link := bridge.LINK;
  END_FOR;
  ASSERT_EQ(ra.ERROR_ID, 1);
  ASSERT_EQ(ra.ABORT_CODE, 16#06020000);
  ASSERT_EQ(rt.ERROR_ID, 2);
  ASSERT_EQ(rt.ABORT_CODE, 16#05040000);
END_TEST

TEST 'bridge gone during a transfer ends with 20'
  VAR
    link : ARRAY[0..1279] OF WORD;
    svc : CW_LINK_SERVICE;
    bridge : MailboxModel;
    rb : CO_SDO_READ_BYTES;
    buf : ARRAY[0..1023] OF BYTE;
  END_VAR
  link[21] := 1;
  link[89] := 16#0431;
  svc(LINK := link);
  rb(EXECUTE := TRUE, NODE := 5, INDEX := 16#2000, BUFFER := buf, LINK := link);
  bridge(LINK := link);
  link := bridge.LINK;
  ASSERT_TRUE(rb.BUSY);
  link[21] := 0;
  svc(LINK := link);
  rb(EXECUTE := TRUE, NODE := 5, INDEX := 16#2000, BUFFER := buf, LINK := link);
  ASSERT_TRUE(rb.ERROR);
  ASSERT_EQ(rb.ERROR_ID, 20);
  ASSERT_EQ(link[94], 0);
END_TEST

TEST 'a waiting instance that is no longer called is skipped'
  VAR
    link : ARRAY[0..1279] OF WORD;
    svc : CW_LINK_SERVICE;
    bridge : MailboxModel;
    s1 : CAN_SEND;
    s2 : CAN_SEND;
    s3 : CAN_SEND;
    d : ARRAY[0..7] OF BYTE;
    i : INT;
  END_VAR
  link[21] := 1;
  link[89] := 16#0431;
  svc(LINK := link);
  s1(EXECUTE := TRUE, ID := 1, DATA := d, LINK := link);
  s2(EXECUTE := TRUE, ID := 2, DATA := d, LINK := link);
  s3(EXECUTE := TRUE, ID := 3, DATA := d, LINK := link);
  bridge(LINK := link);
  link := bridge.LINK;
  (* s2 is never called again *)
  FOR i := 1 TO 8 DO
    svc(LINK := link);
    s1(EXECUTE := TRUE, ID := 1, DATA := d, LINK := link);
    s3(EXECUTE := TRUE, ID := 3, DATA := d, LINK := link);
    bridge(LINK := link);
    link := bridge.LINK;
  END_FOR;
  ASSERT_TRUE(s1.DONE);
  ASSERT_TRUE(s3.DONE);
  ASSERT_EQ(bridge.TX_COUNT, 2);
END_TEST

TEST 'CAN_RECEIVE drains a batch in one scan'
  VAR
    link : ARRAY[0..1279] OF WORD;
    svc : CW_LINK_SERVICE;
    bridge : MailboxModel;
    rx : CAN_RECEIVE;
    d : ARRAY[0..7] OF BYTE;
    i : INT;
    got : INT;
    ids : ARRAY[0..9] OF UDINT;
  END_VAR
  link[21] := 1;
  link[89] := 16#0431;
  FOR i := 1 TO 4 DO
    svc(LINK := link);
    rx(ENABLE := TRUE, ID := 16#180, MASK := 16#780, RX_DATA := d, LINK := link);
    bridge(LINK := link);
    link := bridge.LINK;
  END_FOR;
  ASSERT_TRUE(rx.ACTIVE);
  FOR i := 0 TO 4 DO
    bridge(INJ_CAN := TRUE, INJ_ID := 16#181 + INT_TO_UDINT(i), INJ_DLC := 2, INJ_B0 := INT_TO_BYTE(10 * i), HOLD := TRUE,
           LINK := link);
    link := bridge.LINK;
  END_FOR;
  bridge(INJ_CAN := TRUE, INJ_ID := 16#281, HOLD := FALSE, LINK := link);
  link := bridge.LINK;
  svc(LINK := link);
  rx(ENABLE := TRUE, ID := 16#180, MASK := 16#780, RX_DATA := d, LINK := link);
  WHILE rx.RECEIVED DO
    ids[got] := rx.RX_ID;
    got := got + 1;
    IF got = 5 THEN
      ASSERT_EQ(d[0], 40);
      ASSERT_EQ(d[1], 41);
      ASSERT_EQ(rx.RX_DLC, 2);
    END_IF;
    rx(ENABLE := TRUE, ID := 16#180, MASK := 16#780, RX_DATA := d, LINK := link);
  END_WHILE;
  ASSERT_EQ(got, 5);
  ASSERT_EQ(ids[0], 16#181);
  ASSERT_EQ(ids[4], 16#185);
  ASSERT_EQ(link[104], 0);
  (* acknowledged: the next batch can come *)
  bridge(INJ_CAN := TRUE, INJ_ID := 16#186, LINK := link);
  link := bridge.LINK;
  svc(LINK := link);
  rx(ENABLE := TRUE, ID := 16#180, MASK := 16#780, RX_DATA := d, LINK := link);
  ASSERT_TRUE(rx.RECEIVED);
  ASSERT_EQ(rx.RX_ID, 16#186);
  (* disabled: the receiver closes *)
  FOR i := 1 TO 4 DO
    svc(LINK := link);
    rx(ENABLE := FALSE, RX_DATA := d, LINK := link);
    bridge(LINK := link);
    link := bridge.LINK;
  END_FOR;
  ASSERT_FALSE(rx.ACTIVE);
  ASSERT_EQ(bridge.OPEN_RX, 0);
END_TEST

TEST 'CAN_RECEIVE takes 9 frames a batch with one receive block, all with the batch TIMESTAMP'
  VAR
    link : ARRAY[0..1279] OF WORD;
    svc : CW_LINK_SERVICE;
    bridge : MailboxModel;
    rx : CAN_RECEIVE;
    d : ARRAY[0..7] OF BYTE;
    i : INT;
    got : INT;
    t0 : ULINT;
    same : BOOL;
  END_VAR
  link[21] := 1;
  link[89] := 16#0431;
  FOR i := 1 TO 4 DO
    svc(LINK := link);
    rx(ENABLE := TRUE, ID := 16#180, MASK := 16#780, RX_DATA := d, LINK := link);
    bridge(RX_BLOCKS := 1, LINK := link);
    link := bridge.LINK;
  END_FOR;
  ASSERT_TRUE(rx.ACTIVE);
  FOR i := 0 TO 29 DO
    bridge(INJ_CAN := TRUE, INJ_ID := 16#181, INJ_B0 := INT_TO_BYTE(i), HOLD := TRUE, RX_BLOCKS := 1, LINK := link);
    link := bridge.LINK;
  END_FOR;
  bridge(HOLD := FALSE, RX_BLOCKS := 1, LINK := link);
  link := bridge.LINK;
  svc(LINK := link);
  rx(ENABLE := TRUE, ID := 16#180, MASK := 16#780, RX_DATA := d, LINK := link);
  same := TRUE;
  t0 := rx.TIMESTAMP;
  WHILE rx.RECEIVED DO
    ASSERT_EQ(d[0], INT_TO_BYTE(got));
    same := same AND rx.TIMESTAMP = t0;
    got := got + 1;
    rx(ENABLE := TRUE, ID := 16#180, MASK := 16#780, RX_DATA := d, LINK := link);
  END_WHILE;
  ASSERT_EQ(got, 9);
  ASSERT_TRUE(same);
  (* the next batch: the next frame, with its own time *)
  bridge(RX_BLOCKS := 1, LINK := link);
  link := bridge.LINK;
  svc(LINK := link);
  rx(ENABLE := TRUE, ID := 16#180, MASK := 16#780, RX_DATA := d, LINK := link);
  ASSERT_TRUE(rx.RECEIVED);
  ASSERT_EQ(d[0], INT_TO_BYTE(9));
  ASSERT_TRUE(rx.TIMESTAMP <> t0);
END_TEST

TEST 'CAN_RECEIVE takes 21 frames a batch with two receive blocks'
  VAR
    link : ARRAY[0..1279] OF WORD;
    svc : CW_LINK_SERVICE;
    bridge : MailboxModel;
    rx : CAN_RECEIVE;
    d : ARRAY[0..7] OF BYTE;
    i : INT;
    got : INT;
    t0 : ULINT;
    same : BOOL;
  END_VAR
  link[21] := 1;
  link[89] := 16#0431;
  FOR i := 1 TO 4 DO
    svc(LINK := link);
    rx(ENABLE := TRUE, ID := 16#180, MASK := 16#780, RX_DATA := d, LINK := link);
    bridge(RX_BLOCKS := 2, LINK := link);
    link := bridge.LINK;
  END_FOR;
  ASSERT_TRUE(rx.ACTIVE);
  FOR i := 0 TO 29 DO
    bridge(INJ_CAN := TRUE, INJ_ID := 16#181, INJ_B0 := INT_TO_BYTE(i), HOLD := TRUE, RX_BLOCKS := 2, LINK := link);
    link := bridge.LINK;
  END_FOR;
  bridge(HOLD := FALSE, RX_BLOCKS := 2, LINK := link);
  link := bridge.LINK;
  svc(LINK := link);
  rx(ENABLE := TRUE, ID := 16#180, MASK := 16#780, RX_DATA := d, LINK := link);
  same := TRUE;
  t0 := rx.TIMESTAMP;
  WHILE rx.RECEIVED DO
    ASSERT_EQ(d[0], INT_TO_BYTE(got));
    same := same AND rx.TIMESTAMP = t0;
    got := got + 1;
    rx(ENABLE := TRUE, ID := 16#180, MASK := 16#780, RX_DATA := d, LINK := link);
  END_WHILE;
  ASSERT_EQ(got, 21);
  ASSERT_TRUE(same);
  (* the next batch: the next frame, with its own time *)
  bridge(RX_BLOCKS := 2, LINK := link);
  link := bridge.LINK;
  svc(LINK := link);
  rx(ENABLE := TRUE, ID := 16#180, MASK := 16#780, RX_DATA := d, LINK := link);
  ASSERT_TRUE(rx.RECEIVED);
  ASSERT_EQ(d[0], INT_TO_BYTE(21));
  ASSERT_TRUE(rx.TIMESTAMP <> t0);
END_TEST

TEST 'CAN_RECEIVE keeps receiving as the bridge clock wraps'
  VAR
    link : ARRAY[0..1279] OF WORD;
    svc : CW_LINK_SERVICE;
    bridge : MailboxModel;
    rx : CAN_RECEIVE;
    d : ARRAY[0..7] OF BYTE;
    i : INT;
    k : INT;
    got : INT;
  END_VAR
  link[21] := 1;
  link[89] := 16#0431;
  FOR i := 1 TO 4 DO
    svc(LINK := link);
    rx(ENABLE := TRUE, ID := 16#180, MASK := 16#780, RX_DATA := d, LINK := link);
    bridge(LINK := link);
    link := bridge.LINK;
  END_FOR;
  ASSERT_TRUE(rx.ACTIVE);
  (* one frame every 10 s of bridge time, for more than one 65.5 s wrap *)
  FOR k := 1 TO 10 DO
    bridge(INJ_CAN := TRUE, INJ_ID := 16#181, SKIP_MS := 10000, LINK := link);
    link := bridge.LINK;
    svc(LINK := link);
    rx(ENABLE := TRUE, ID := 16#180, MASK := 16#780, RX_DATA := d, LINK := link);
    IF rx.RECEIVED THEN
      got := got + 1;
      rx(ENABLE := TRUE, ID := 16#180, MASK := 16#780, RX_DATA := d, LINK := link);
    END_IF;
  END_FOR;
  ASSERT_EQ(got, 10);
  ASSERT_TRUE(rx.ACTIVE);
  ASSERT_FALSE(rx.ERROR);
END_TEST

TEST 'a receiver the bridge closed opens again'
  VAR
    link : ARRAY[0..1279] OF WORD;
    svc : CW_LINK_SERVICE;
    bridge : MailboxModel;
    rx : CAN_RECEIVE;
    d : ARRAY[0..7] OF BYTE;
    i : INT;
    saw8 : BOOL;
  END_VAR
  link[21] := 1;
  link[89] := 16#0431;
  FOR i := 1 TO 4 DO
    svc(LINK := link);
    rx(ENABLE := TRUE, ID := 16#180, RX_DATA := d, LINK := link);
    bridge(LINK := link);
    link := bridge.LINK;
  END_FOR;
  ASSERT_TRUE(rx.ACTIVE);
  bridge(CLOSE_SLOT := 0, LINK := link);
  link := bridge.LINK;
  FOR i := 1 TO 6 DO
    svc(LINK := link);
    rx(ENABLE := TRUE, ID := 16#180, RX_DATA := d, LINK := link);
    IF rx.ERROR_ID = 8 THEN
      saw8 := TRUE;
    END_IF;
    bridge(LINK := link);
    link := bridge.LINK;
  END_FOR;
  ASSERT_TRUE(saw8);
  ASSERT_TRUE(rx.ACTIVE);
  ASSERT_FALSE(rx.ERROR);
END_TEST

TEST 'CAN_SEND_CYCLIC starts, updates only on change and stops'
  VAR
    link : ARRAY[0..1279] OF WORD;
    svc : CW_LINK_SERVICE;
    bridge : MailboxModel;
    cyc : CAN_SEND_CYCLIC;
    d : ARRAY[0..7] OF BYTE;
    i : INT;
  END_VAR
  link[21] := 1;
  link[89] := 16#0431;
  d[0] := 1;
  FOR i := 1 TO 10 DO
    svc(LINK := link);
    cyc(ENABLE := TRUE, ID := 16#200, DLC := 1, PERIOD := T#20ms, DATA := d, LINK := link);
    bridge(LINK := link);
    link := bridge.LINK;
  END_FOR;
  ASSERT_TRUE(cyc.ACTIVE);
  ASSERT_EQ(bridge.CYC_SETS, 1);
  ASSERT_TRUE(cyc.COUNT > 3);
  d[0] := 2;
  FOR i := 1 TO 5 DO
    svc(LINK := link);
    cyc(ENABLE := TRUE, ID := 16#200, DLC := 1, PERIOD := T#20ms, DATA := d, LINK := link);
    bridge(LINK := link);
    link := bridge.LINK;
  END_FOR;
  ASSERT_EQ(bridge.CYC_SETS, 2);
  ASSERT_EQ(bridge.job_data[0], 16#0200);
  FOR i := 1 TO 5 DO
    svc(LINK := link);
    cyc(ENABLE := FALSE, DATA := d, LINK := link);
    bridge(LINK := link);
    link := bridge.LINK;
  END_FOR;
  ASSERT_FALSE(cyc.ACTIVE);
  ASSERT_EQ(bridge.CYC_STOPS, 1);
  ASSERT_FALSE(bridge.job_on[0]);
END_TEST

TEST 'bus info and ECU info from the info block'
  VAR
    link : ARRAY[0..1279] OF WORD;
    bridge : MailboxModel;
    bus : CAN_BUS_INFO;
    ecu : J1939_ECU_INFO;
    other : J1939_ECU_INFO;
  END_VAR
  link[21] := 1;
  link[89] := 16#0431;
  bridge(LINK := link);
  link := bridge.LINK;
  bus(NETWORK := 0, LINK := link);
  ASSERT_FALSE(bus.ERROR);
  ASSERT_EQ(bus.STATE, 0);
  ASSERT_EQ(bus.BUS_LOAD, 12);
  ASSERT_EQ(bus.BUS_OFF_COUNT, 3);
  ASSERT_EQ(bus.RX_COUNT, 1000);
  ASSERT_EQ(bus.TX_COUNT, 65536);
  ecu(ENABLE := TRUE, NETWORK := 0, LINK := link);
  ASSERT_TRUE(ecu.VALID);
  ASSERT_EQ(ecu.STATE, 1);
  ASSERT_EQ(ecu.ADDRESS, 16#80);
  ASSERT_EQ(ecu.NAME, 16#A00000000000ABCD);
  ASSERT_EQ(ecu.ECU_COUNT, 4);
  other(ENABLE := TRUE, NETWORK := 1, LINK := link);
  ASSERT_EQ(other.ERROR_ID, 10);
  bus(NETWORK := 2, LINK := link);
  ASSERT_EQ(bus.ERROR_ID, 2);
END_TEST

TEST 'J1939 send short and long, request long, DM read and clear, find ECU'
  VAR
    link : ARRAY[0..1279] OF WORD;
    svc : CW_LINK_SERVICE;
    bridge : MailboxModel;
    snd : J1939_SEND;
    req : J1939_REQUEST;
    nack : J1939_REQUEST;
    dm : J1939_DM_READ;
    clr : J1939_DM_CLEAR;
    find : J1939_FIND_ECU;
    data : ARRAY[0..1784] OF BYTE;
    rdata : ARRAY[0..1784] OF BYTE;
    ndata : ARRAY[0..1784] OF BYTE;
    dtcs : ARRAY[0..31] OF UDINT;
    i : INT;
  END_VAR
  link[21] := 1;
  link[89] := 16#0431;
  FOR i := 0 TO 299 DO
    data[i] := INT_TO_BYTE(i MOD 13);
  END_FOR;
  FOR i := 1 TO 40 DO
    svc(LINK := link);
    snd(EXECUTE := TRUE, PGN := 65281, DESTINATION := 255, LENGTH := 300, DATA := data, LINK := link);
    req(EXECUTE := TRUE, PGN := 65000, DESTINATION := 16#21, DATA := rdata, LINK := link);
    nack(EXECUTE := TRUE, PGN := 59999, DESTINATION := 16#21, DATA := ndata, LINK := link);
    dm(EXECUTE := TRUE, SOURCE := 0, DTCS := dtcs, LINK := link);
    clr(EXECUTE := TRUE, DESTINATION := 9, LINK := link);
    find(ENABLE := TRUE, NAME := 16#A000000000000000, MASK := 16#FF00000000000000, LINK := link);
    bridge(LINK := link);
    link := bridge.LINK;
  END_FOR;
  ASSERT_TRUE(snd.DONE);
  ASSERT_EQ(bridge.J_LEN, 300);
  ASSERT_EQ(bridge.J_PRIO, 6);
  ASSERT_EQ(bridge.j_data[299], 0);
  ASSERT_EQ(bridge.j_data[140], 10);
  ASSERT_TRUE(req.DONE);
  ASSERT_EQ(req.LENGTH, 300);
  ASSERT_EQ(req.SOURCE, 16#21);
  ASSERT_EQ(rdata[299], 43);
  ASSERT_TRUE(nack.ERROR);
  ASSERT_EQ(nack.ERROR_ID, 12);
  ASSERT_EQ(nack.ACK_CODE, 1);
  ASSERT_TRUE(dm.DONE);
  ASSERT_EQ(dm.COUNT, 2);
  ASSERT_EQ(dm.LAMPS, 16#44);
  ASSERT_EQ(dm.FLASH, 16#04);
  ASSERT_EQ(dm.AGE, T#1500ms);
  ASSERT_EQ(dtcs[0], 16#00012304);
  ASSERT_EQ(dtcs[1], 16#0005A1FF);
  ASSERT_TRUE(clr.DONE);
  ASSERT_EQ(bridge.DM_CLEARED, 9);
  ASSERT_TRUE(find.VALID);
  ASSERT_TRUE(find.FOUND);
  ASSERT_EQ(find.ADDRESS, 16#33);
  ASSERT_EQ(find.FOUND_NAME, 16#A00000000000ABCD);
END_TEST

TEST 'J1939_RECEIVE reads a long message whole'
  VAR
    link : ARRAY[0..1279] OF WORD;
    svc : CW_LINK_SERVICE;
    bridge : MailboxModel;
    rx : J1939_RECEIVE;
    data : ARRAY[0..1784] OF BYTE;
    i : INT;
    got : BOOL;
  END_VAR
  link[21] := 1;
  link[89] := 16#0431;
  FOR i := 1 TO 4 DO
    svc(LINK := link);
    rx(ENABLE := TRUE, PGN := 65282, RX_DATA := data, LINK := link);
    bridge(LINK := link);
    link := bridge.LINK;
  END_FOR;
  ASSERT_TRUE(rx.ACTIVE);
  bridge(INJ_J1939 := TRUE, INJ_ID := 65282, INJ_LEN := 200, INJ_SRC := 0, INJ_B0 := 1, LINK := link);
  link := bridge.LINK;
  FOR i := 1 TO 10 DO
    svc(LINK := link);
    rx(ENABLE := TRUE, PGN := 65282, RX_DATA := data, LINK := link);
    IF rx.RECEIVED THEN
      got := TRUE;
      ASSERT_EQ(rx.RX_LENGTH, 200);
      ASSERT_EQ(rx.RX_PGN, 65282);
      ASSERT_EQ(data[0], 1);
      ASSERT_EQ(data[199], 200);
    END_IF;
    bridge(LINK := link);
    link := bridge.LINK;
  END_FOR;
  ASSERT_TRUE(got);
  ASSERT_FALSE(rx.ERROR);
END_TEST

TEST 'two EMCY receivers each get a message; a new session shows 8 once'
  VAR
    link : ARRAY[0..1279] OF WORD;
    svc : CW_LINK_SERVICE;
    bridge : MailboxModel;
    e1 : CO_RECV_EMCY;
    e2 : CO_RECV_EMCY;
    m1 : ARRAY[0..4] OF BYTE;
    m2 : ARRAY[0..4] OF BYTE;
    i : INT;
    n1 : INT;
    n2 : INT;
    eights : INT;
  END_VAR
  link[21] := 1;
  link[89] := 16#0431;
  FOR i := 1 TO 6 DO
    svc(LINK := link);
    e1(ENABLE := TRUE, MSEF := m1, LINK := link);
    e2(ENABLE := TRUE, NODE := 3, MSEF := m2, LINK := link);
    bridge(LINK := link);
    link := bridge.LINK;
  END_FOR;
  ASSERT_TRUE(e1.ACTIVE);
  ASSERT_TRUE(e2.ACTIVE);
  bridge(INJ_EMCY := TRUE, INJ_NODE := 3, INJ_CODE := 16#8130, LINK := link);
  link := bridge.LINK;
  FOR i := 1 TO 4 DO
    svc(LINK := link);
    e1(ENABLE := TRUE, MSEF := m1, LINK := link);
    e2(ENABLE := TRUE, NODE := 3, MSEF := m2, LINK := link);
    IF e1.RECEIVED THEN
      n1 := n1 + 1;
      ASSERT_EQ(e1.ERROR_CODE, 16#8130);
      ASSERT_EQ(e1.EMCY_NODE, 3);
      ASSERT_EQ(e1.ERROR_REGISTER, 16#81);
      ASSERT_EQ(m1[4], 5);
    END_IF;
    IF e2.RECEIVED THEN
      n2 := n2 + 1;
    END_IF;
    bridge(LINK := link);
    link := bridge.LINK;
  END_FOR;
  ASSERT_EQ(n1, 1);
  ASSERT_EQ(n2, 1);
  bridge(INJ_RESTART := TRUE, INJ_NODE := 3, LINK := link);
  link := bridge.LINK;
  FOR i := 1 TO 4 DO
    svc(LINK := link);
    e1(ENABLE := TRUE, MSEF := m1, LINK := link);
    IF e1.ERROR_ID = 8 THEN
      eights := eights + 1;
    END_IF;
    bridge(LINK := link);
    link := bridge.LINK;
  END_FOR;
  ASSERT_EQ(eights, 1);
  ASSERT_TRUE(e1.ACTIVE);
END_TEST

(* ---- test_programs.st ---- *)
(*
 * The generated canworks_in and canworks_out (tools/deploy/canworks/
 * openplcmodbus.py) for test/plc_modbus/canworks.json, as function blocks
 * (make_programs.py): raw Modbus words to typed values and back, low word
 * first, and the PLC link header. Run by test/plc_modbus/run.sh.
 *)
TEST 'canworks_in converts the input registers'
  VAR
    cin : canworks_in_fb;
  END_VAR
  cin.i0 := 16#EC2C;
  cin.i1 := 16#168F;
  cin.i3 := 5;
  cin.i6 := 16#0380;
  cin.i7 := 16#FF05;
  cin.i8 := 16#FFFE;
  cin.i9 := 16#7960;
  cin.i10 := 16#FFFE;
  cin.i11 := 16#0000;
  cin.i12 := 16#3FC0;
  cin.i13 := 16#CDEF;
  cin.i14 := 16#89AB;
  cin.i15 := 16#4567;
  cin.i16 := 16#0123;
  cin.i17 := 0;
  cin.i18 := 0;
  cin.i19 := 0;
  cin.i20 := 16#C004;
  cin.i21 := 7;
  cin();
  ASSERT_TRUE(cin.canworks.ok);
  ASSERT_EQ(cin.canworks.link[21], 16#0007);
  ASSERT_TRUE(cin.canworks.cab_In_status);
  ASSERT_TRUE(cin.canworks.cab_In_flag);
  ASSERT_TRUE(cin.canworks.cab_In_low);
  ASSERT_EQ(cin.canworks.cab_In_sbyte, -1);
  ASSERT_EQ(cin.canworks.cab_In_ubyte, 5);
  ASSERT_EQ(cin.canworks.cab_In_word, -2);
  ASSERT_EQ(cin.canworks.cab_In_dword, -100000);
  ASSERT_NEAR(cin.canworks.cab_In_real, 1.5, 0.0);
  ASSERT_EQ(cin.canworks.cab_Wide_lword, ULINT#16#0123456789ABCDEF);
  ASSERT_NEAR(cin.canworks.cab_Wide_lreal, -2.5, 0.0);
  ASSERT_EQ(cin.canworks.link[14], 7);
END_TEST

TEST 'canworks.ok needs the map hash and a moving counter'
  VAR
    cin : canworks_in_fb;
  END_VAR
  cin.i0 := 16#EC2C;
  cin.i1 := 16#1690;
  cin.i3 := 1;
  cin();
  ASSERT_FALSE(cin.canworks.ok);
  cin.i1 := 16#168F;
  cin.i3 := 2;
  cin();
  ASSERT_TRUE(cin.canworks.ok);
  cin();
  ADVANCE_TIME(T#200ms);
  cin();
  ASSERT_TRUE(cin.canworks.ok);
  ADVANCE_TIME(T#200ms);
  cin();
  ASSERT_FALSE(cin.canworks.ok);
  cin.i3 := 3;
  cin();
  ASSERT_TRUE(cin.canworks.ok);
  cin.i0 := 0;
  cin.i1 := 0;
  cin.i3 := 4;
  cin();
  ASSERT_FALSE(cin.canworks.ok);
END_TEST

TEST 'while canworks.ok is FALSE the status inputs read 0 and the others hold'
  VAR
    cin : canworks_in_fb;
  END_VAR
  cin.i0 := 16#EC2C;
  cin.i1 := 16#168F;
  cin.i3 := 1;
  cin.i6 := 16#0300;
  cin.i8 := 16#FFFE;
  cin();
  ASSERT_TRUE(cin.canworks.ok);
  ASSERT_TRUE(cin.canworks.bus_ok);
  ASSERT_TRUE(cin.canworks.cab_In_status);
  ASSERT_TRUE(cin.canworks.cab_In_flag);
  ASSERT_EQ(cin.canworks.cab_In_word, -2);
  (* The counter stops: the bridge is lost. *)
  cin();
  ADVANCE_TIME(T#400ms);
  cin();
  ASSERT_FALSE(cin.canworks.ok);
  ASSERT_FALSE(cin.canworks.bus_ok);
  ASSERT_FALSE(cin.canworks.cab_In_status);
  ASSERT_TRUE(cin.canworks.cab_In_flag);
  ASSERT_EQ(cin.canworks.cab_In_word, -2);
END_TEST

TEST 'inputs_on_loss zero sets every input to 0 while canworks.ok is FALSE'
  VAR
    cin : canworks_in_zero_fb;
  END_VAR
  cin.i0 := 16#EC2C;
  cin.i1 := 16#168F;
  cin.i3 := 1;
  cin.i6 := 16#0300;
  cin.i8 := 16#FFFE;
  cin.i11 := 16#0000;
  cin.i12 := 16#3FC0;
  cin();
  ASSERT_TRUE(cin.canworks.cab_In_flag);
  ASSERT_EQ(cin.canworks.cab_In_word, -2);
  ASSERT_NEAR(cin.canworks.cab_In_real, 1.5, 0.0);
  cin();
  ADVANCE_TIME(T#400ms);
  cin();
  ASSERT_FALSE(cin.canworks.ok);
  ASSERT_FALSE(cin.canworks.cab_In_status);
  ASSERT_FALSE(cin.canworks.cab_In_flag);
  ASSERT_EQ(cin.canworks.cab_In_word, 0);
  ASSERT_NEAR(cin.canworks.cab_In_real, 0.0, 0.0);
END_TEST

TEST 'canworks.bus_ok follows status byte 7 bit 1'
  VAR
    cin : canworks_in_fb;
  END_VAR
  cin.i0 := 16#EC2C;
  cin.i1 := 16#168F;
  cin.i3 := 1;
  cin.i5 := 16#0002;
  cin();
  ASSERT_TRUE(cin.canworks.ok);
  ASSERT_FALSE(cin.canworks.bus_ok);
  cin.i3 := 2;
  cin.i5 := 16#0001;
  cin();
  ASSERT_TRUE(cin.canworks.bus_ok);
END_TEST

TEST 'canworks_out writes the holding registers and the header last'
  VAR
    cout : canworks_out_fb;
  END_VAR
  cout.canworks.cab_Out_flag := TRUE;
  cout.canworks.cab_Out_low := TRUE;
  cout.canworks.cab_Out_sbyte := -2;
  cout.canworks.cab_Out_ubyte := 7;
  cout.canworks.cab_Out_word := -3;
  cout.canworks.cab_Out_dword := -100000;
  cout.canworks.cab_Out_real := 1.5;
  cout.canworks.cab_Wide_lreal_2 := -2.5;
  cout.canworks.link[5] := 16#0400;
  cout.canworks.link[13] := 16#BEEF;
  cout();
  ASSERT_EQ(cout.q0, 1);
  ASSERT_EQ(cout.q1, 16#EC2C);
  ASSERT_EQ(cout.q2, 16#168F);
  ASSERT_EQ(cout.q3, 16#0108);
  ASSERT_EQ(cout.q4, 16#FE07);
  ASSERT_EQ(cout.q5, 16#FFFD);
  ASSERT_EQ(cout.q6, 16#7960);
  ASSERT_EQ(cout.q7, 16#FFFE);
  ASSERT_EQ(cout.q8, 16#0000);
  ASSERT_EQ(cout.q9, 16#3FC0);
  ASSERT_EQ(cout.q10, 0);
  ASSERT_EQ(cout.q13, 16#C004);
  ASSERT_EQ(cout.q15, 16#0400);
  ASSERT_EQ(cout.q23, 16#BEEF);
END_TEST

TEST 'mailbox words go between the registers and LINK, the link service runs'
  VAR
    cin : canworks_in_fb;
    cout : canworks_out_fb;
  END_VAR
  (* responses from input register 28, the receive mailbox from 100, info
     from 220, the cyclic table from 238; requests from holding register 24,
     the acknowledgement from 96, keepalives from 99 *)
  cin.i0 := 16#EC2C;
  cin.i1 := 16#168F;
  cin.i3 := 1;
  cin.i28 := 16#0042;
  cin.i99 := 16#5A5A;
  cin.i100 := 16#7001;
  cin.i220 := 16#000C;
  cin.i254 := 16#0009;
  cin();
  ASSERT_EQ(cin.canworks.link[89], 16#0431);
  ASSERT_EQ(cin.canworks.link[216], 16#0042);
  ASSERT_EQ(cin.canworks.link[287], 16#5A5A);
  ASSERT_EQ(cin.canworks.link[720], 16#7001);
  ASSERT_EQ(cin.canworks.link[960], 16#000C);
  ASSERT_EQ(cin.canworks.link[1120], 16#0009);
  (* CW_LINK_SERVICE ran: one scan, the new batch acknowledged *)
  ASSERT_EQ(cin.canworks.link[90], 1);
  ASSERT_EQ(cin.canworks.link[102], 16#7001);
  cout.canworks.link[144] := 16#0101;
  cout.canworks.link[215] := 16#0202;
  cout.canworks.link[102] := 16#7001;
  cout.canworks.link[131] := 16#0303;
  cout();
  ASSERT_EQ(cout.q24, 16#0101);
  ASSERT_EQ(cout.q95, 16#0202);
  ASSERT_EQ(cout.q96, 16#7001);
  ASSERT_EQ(cout.q102, 16#0303);
END_TEST
